(* IEC 61131-3 sources: model-first-plc-agent-ai/results/T4-W-08, 2 files *)

(* ---- a1_code.st ---- *)
FUNCTION_BLOCK LevelControlRuntime
VAR_INPUT
    StartSignal : BOOL;
    StopSignal : BOOL;
    LevelValue : INT;
    FullScaleValue : INT;
    h_span : REAL;
    h_target : REAL;
    h_sp : REAL;
    h_max : REAL;
    eps : REAL;
    t_h : TIME;
    Kp : REAL;
    Ti : REAL;
    Td : REAL;
    CycleSeconds : REAL;
END_VAR
VAR_OUTPUT
    fill_valve : BOOL;
    discharge_valve : BOOL;
    FillCommand : INT;
    DischargeCommand : INT;
END_VAR
VAR
    StartEdge : R_TRIG;
    HoldTimer : TON;
    start : BOOL;
    stop : BOOL;
    settled : BOOL;
    r : INT;
    x0 : BOOL := TRUE;
    x1 : BOOL := FALSE;
    ActiveState : INT := 0;
    h : REAL;
    ErrorValue : REAL;
    PreviousError : REAL := 0.0;
    DerivativeReady : BOOL := FALSE;
    ProportionalTerm : REAL;
    IntegralTerm : REAL := 0.0;
    CandidateIntegral : REAL;
    DerivativeTerm : REAL;
    RawDemand : REAL;
    CandidateDemand : REAL;
    BoundedDemand : REAL;
END_VAR
VAR CONSTANT
    RegionLow : INT := 0;
    RegionMiddle : INT := 1;
    RegionHigh : INT := 2;
END_VAR

StartEdge(CLK := StartSignal);
start := StartEdge.Q;
stop := StopSignal;

h := INT_TO_REAL(LevelValue) * h_span / INT_TO_REAL(FullScaleValue);
ErrorValue := h_sp - h;

IF h < h_target THEN
    r := RegionLow;
ELSIF h < h_max THEN
    r := RegionMiddle;
ELSE
    r := RegionHigh;
END_IF;

(* The tolerance interval must remain continuous during step x1. *)
HoldTimer(
    IN := x1 AND NOT stop AND (ABS(ErrorValue) <= eps),
    PT := t_h
);
settled := HoldTimer.Q;

(* Evaluate transitions from the situation at the start of this scan. *)
CASE ActiveState OF
    0:
        IF start AND NOT stop AND (r <> RegionHigh) THEN
            ActiveState := 1;
        END_IF;

    1:
        IF stop OR settled OR (r = RegionHigh) THEN
            ActiveState := 0;
        END_IF;
ELSE
    ActiveState := 0;
END_CASE;

x0 := ActiveState = 0;
x1 := ActiveState = 1;

fill_valve := x1;
discharge_valve := x1;

FillCommand := 0;
DischargeCommand := 0;

IF fill_valve THEN
    (* Parallel PID, with demand expressed as percent valve opening.
       Ti and Td are in seconds; Kp is percent opening per level unit. *)
    ProportionalTerm := Kp * ErrorValue;
    DerivativeTerm := 0.0;

    IF DerivativeReady AND (CycleSeconds > 0.0) THEN
        DerivativeTerm :=
            Kp * Td * (ErrorValue - PreviousError) / CycleSeconds;
    END_IF;

    RawDemand := ProportionalTerm + IntegralTerm + DerivativeTerm;
    CandidateIntegral := IntegralTerm;

    IF (Ti > 0.0) AND (CycleSeconds > 0.0) THEN
        CandidateIntegral :=
            IntegralTerm + Kp * ErrorValue * CycleSeconds / Ti;
    END_IF;

    CandidateDemand :=
        ProportionalTerm + CandidateIntegral + DerivativeTerm;

    (* Freeze integration whenever the output is clamped.
       Also reject an integral update that would cause clamping. *)
    IF (RawDemand >= 0.0) AND (RawDemand <= 100.0)
        AND (CandidateDemand >= 0.0)
        AND (CandidateDemand <= 100.0) THEN
        IntegralTerm := CandidateIntegral;
    END_IF;

    RawDemand := ProportionalTerm + IntegralTerm + DerivativeTerm;

    IF RawDemand > 100.0 THEN
        BoundedDemand := 100.0;
    ELSIF RawDemand < 0.0 THEN
        BoundedDemand := 0.0;
    ELSE
        BoundedDemand := RawDemand;
    END_IF;

    FillCommand :=
        REAL_TO_INT(BoundedDemand * INT_TO_REAL(FullScaleValue) / 100.0);

    PreviousError := ErrorValue;
    DerivativeReady := TRUE;
ELSE
    (* No stored action: the idle step explicitly closes both valves. *)
    IntegralTerm := 0.0;
    PreviousError := ErrorValue;
    DerivativeReady := FALSE;
    BoundedDemand := 0.0;
END_IF;

IF discharge_valve THEN
    DischargeCommand := REAL_TO_INT(0.4 * INT_TO_REAL(FullScaleValue));
END_IF;

END_FUNCTION_BLOCK

PROGRAM Main
VAR
    StartCommand AT %IX100.0 : BOOL;
    StopCommand AT %IX100.1 : BOOL;
    LevelMeter AT %IW100 : INT;
    FillValve AT %QW100 : INT;
    DischargeValve AT %QW101 : INT;
END_VAR
VAR CONSTANT
    FULL_SCALE : INT := 1000;
END_VAR
VAR
    Controller : LevelControlRuntime;
    Initialized : BOOL := FALSE;

    h_span : REAL := 10.0;
    h_target : REAL;
    h_sp : REAL;
    h_max : REAL;
    eps : REAL;
    t_h : TIME := T#10s;

    (* Commissioning parameters; tune for the simulated plant. *)
    Kp : REAL := 10.0;
    Ti : REAL := 5.0;
    Td : REAL := 0.0;
    CycleSeconds : REAL := 0.02;
END_VAR

IF NOT Initialized THEN
    FillValve := 0;
    DischargeValve := 0;
    Initialized := TRUE;
END_IF;

h_target := 0.8 * h_span;
h_sp := h_target;
h_max := 0.9 * h_span;
eps := 0.02 * h_span;

Controller(
    StartSignal := StartCommand,
    StopSignal := StopCommand,
    LevelValue := LevelMeter,
    FullScaleValue := FULL_SCALE,
    h_span := h_span,
    h_target := h_target,
    h_sp := h_sp,
    h_max := h_max,
    eps := eps,
    t_h := t_h,
    Kp := Kp,
    Ti := Ti,
    Td := Td,
    CycleSeconds := CycleSeconds
);

FillValve := Controller.FillCommand;
DischargeValve := Controller.DischargeCommand;

END_PROGRAM

CONFIGURATION Config0
    RESOURCE Res0 ON PLC
        TASK MainTask(INTERVAL := T#20ms, PRIORITY := 0);
        PROGRAM MainInstance WITH MainTask : Main;
    END_RESOURCE
END_CONFIGURATION

(* ---- a2_code.st ---- *)
FUNCTION_BLOCK FB_LevelControl
VAR_INPUT
    StartCommand : BOOL;
    StopCommand : BOOL;
    LevelMeter : INT;
    h_span : REAL;
    h_target : REAL;
    h_max : REAL;
    eps : REAL;
    t_h : TIME;
    Kp : REAL;
    Ti : REAL;
    Td : REAL;
    CycleSeconds : REAL;
END_VAR
VAR_OUTPUT
    FillValve : INT;
    DischargeValve : INT;
    fill_valve : BOOL;
    discharge_valve : BOOL;
END_VAR
VAR CONSTANT
    FULL_SCALE : INT := 1000;
    REGION_LOW : INT := 0;
    REGION_MIDDLE : INT := 1;
    REGION_HIGH : INT := 2;
END_VAR
VAR
    StartEdge : R_TRIG;
    HoldTimer : TON;
    start : BOOL;
    stop : BOOL;
    settled : BOOL;
    r : INT;
    x0 : BOOL := TRUE;
    x1 : BOOL := FALSE;
    SequenceState : INT := 0;
    WasRegulating : BOOL := FALSE;
    h : REAL;
    h_sp : REAL;
    e : REAL;
    NormalizedError : REAL;
    PreviousError : REAL := 0.0;
    IntegralTerm : REAL := 0.0;
    IntegralCandidate : REAL;
    ProportionalTerm : REAL;
    DerivativeTerm : REAL;
    CandidateDemand : REAL;
    RawDemand : REAL;
    BoundedDemand : REAL;
    ParametersValid : BOOL;
END_VAR

StartEdge(CLK := StartCommand);
start := StartEdge.Q;
stop := StopCommand;

h := INT_TO_REAL(LevelMeter) * h_span / INT_TO_REAL(FULL_SCALE);
h_sp := h_target;
e := h_sp - h;

IF h < h_target THEN
    r := REGION_LOW;
ELSIF h < h_max THEN
    r := REGION_MIDDLE;
ELSE
    r := REGION_HIGH;
END_IF;

ParametersValid :=
    (h_span > 0.0) AND
    (CycleSeconds > 0.0) AND
    (Ti >= 0.0) AND
    (Td >= 0.0);

(* The hold interval measures continuous time inside the tolerance band,
   and is reset whenever regulation is inactive or the band is left. *)
HoldTimer(
    IN := x1 AND NOT stop AND ParametersValid AND (ABS(e) <= eps),
    PT := t_h
);
settled := HoldTimer.Q;

(* Stop has priority over every transition and action. *)
IF stop OR NOT ParametersValid THEN
    SequenceState := 0;
ELSE
    CASE SequenceState OF
        0:
            IF start AND (r <> REGION_HIGH) THEN
                SequenceState := 1;
            END_IF;
        1:
            IF settled OR (r = REGION_HIGH) THEN
                SequenceState := 0;
            END_IF;
    ELSE
        SequenceState := 0;
    END_CASE;
END_IF;

x0 := SequenceState = 0;
x1 := SequenceState = 1;
fill_valve := x1;
discharge_valve := x1;

FillValve := 0;
DischargeValve := 0;

IF x1 THEN
    NormalizedError := e / h_span;

    IF NOT WasRegulating THEN
        IntegralTerm := 0.0;
        PreviousError := NormalizedError;
    END_IF;

    (* Parallel terms implement Kp * (e + integral(e)/Ti + Td*de/dt),
       using error normalized to the measuring span. *)
    ProportionalTerm := Kp * NormalizedError;
    DerivativeTerm :=
        Kp * Td * (NormalizedError - PreviousError) / CycleSeconds;

    IF Ti > 0.0 THEN
        IntegralCandidate :=
            IntegralTerm + Kp * NormalizedError * CycleSeconds / Ti;
    ELSE
        (* Ti = 0 disables integral action. *)
        IntegralTerm := 0.0;
        IntegralCandidate := 0.0;
    END_IF;

    RawDemand := ProportionalTerm + IntegralTerm + DerivativeTerm;
    CandidateDemand :=
        ProportionalTerm + IntegralCandidate + DerivativeTerm;

    (* Suspend integration when the existing or proposed demand is clamped. *)
    IF (RawDemand >= 0.0) AND (RawDemand <= 1.0) AND
       (CandidateDemand >= 0.0) AND (CandidateDemand <= 1.0) THEN
        IntegralTerm := IntegralCandidate;
    END_IF;

    RawDemand := ProportionalTerm + IntegralTerm + DerivativeTerm;

    IF RawDemand < 0.0 THEN
        BoundedDemand := 0.0;
    ELSIF RawDemand > 1.0 THEN
        BoundedDemand := 1.0;
    ELSE
        BoundedDemand := RawDemand;
    END_IF;

    FillValve := REAL_TO_INT(BoundedDemand * INT_TO_REAL(FULL_SCALE));
    DischargeValve := REAL_TO_INT(0.4 * INT_TO_REAL(FULL_SCALE));
    PreviousError := NormalizedError;
ELSE
    IntegralTerm := 0.0;
    PreviousError := 0.0;
    BoundedDemand := 0.0;
END_IF;

WasRegulating := x1;
END_FUNCTION_BLOCK

PROGRAM Main
VAR
    StartCommand AT %IX100.0 : BOOL;
    StopCommand AT %IX100.1 : BOOL;
    LevelMeter AT %IW100 : INT;
    FillValve AT %QW100 : INT;
    DischargeValve AT %QW101 : INT;
END_VAR
VAR
    LevelController : FB_LevelControl;
    fill_valve : BOOL;
    discharge_valve : BOOL;

    h_span : REAL := 10.0;
    h_target : REAL;
    h_max : REAL;
    eps : REAL;
    t_h : TIME := T#10s;

    (* Initial tuning values; adjust for the simulated plant. *)
    Kp : REAL := 1.0;
    Ti : REAL := 10.0;
    Td : REAL := 0.0;

    (* Configure the OpenPLC task to execute Main every 20 ms,
       or change this value to match its actual execution interval. *)
    CycleSeconds : REAL := 0.02;
END_VAR

h_target := 0.8 * h_span;
h_max := 0.9 * h_span;
eps := 0.02 * h_span;

LevelController(
    StartCommand := StartCommand,
    StopCommand := StopCommand,
    LevelMeter := LevelMeter,
    h_span := h_span,
    h_target := h_target,
    h_max := h_max,
    eps := eps,
    t_h := t_h,
    Kp := Kp,
    Ti := Ti,
    Td := Td,
    CycleSeconds := CycleSeconds
);

FillValve := LevelController.FillValve;
DischargeValve := LevelController.DischargeValve;
fill_valve := LevelController.fill_valve;
discharge_valve := LevelController.discharge_valve;
END_PROGRAM
